(* IEC 61131-3 sources: trust-platform/conformance/cases/init_reset/cfm_init_reset_var_initialization_001, 1 file *)

(* ---- program.st ---- *)
PROGRAM Main
VAR
    a : INT;
    b : INT := 4;
    c : INT := b + 1;
END_VAR
END_PROGRAM
